Fanuc KAREL source: IO0225.KL

PROGRAM IO0225
%NOLOCKGROUP
ROUTINE RTEST
VAR
  I : INTEGER
  STATUS : INTEGER
  ENTRY : INTEGER
  A : ARRAY[3] OF INTEGER
  B : BOOLEAN
  R : REAL
  P : XYZWPR
  JPOS : JOINTPOS
  PF : POSITION
BEGIN
  I = 1
  A[1] = 2
  B = TRUE
  R = 1.0
  GET_VAR(ENTRY,'*POSREG*','$MAXPREGNUM',I,STATUS)
END RTEST
BEGIN
  RTEST
END IO0225
